FUNCTION_BLOCK FB_DatamanScanner
(*

The function block used to control scanner.

Constructor: 		Patryk Panylo
Company:		E. Riexinger GmbH
Date:			24.01.2019
Version:			1.00

Date:			Revision:		Who:				Comment
dd.mm.yyyy		x.xx			Initials			comment

*)
VAR_INPUT
	(* Input variables / Eingang Variablen *)
	sSrvNetID				:T_AmsNetID	:= '';						(* TwinCAT TCP/IP server network address *)
	sRemoteHost				:T_IPv4Addr := '192.168.10.1';			(* Server network address *)
	nRemotePort				:UDINT := 23;							(* Server port number *)
	bEnable					:BOOL := FALSE;							(* TRUE => enable client data exchange, FALSE => disable *)
	bReset					:BOOL := FALSE;							(* Confirm alarm *)
	bExecute 				:BOOL := FALSE;							(* Send execute command *)
	bLoggerEn				:BOOL := FALSE;							(* TRUE => Enable log message output, FALSE => Disable *)
	sSndMsg					:T_MaxString := 'BEEP 2 2';				(* Send command is an ASCII typable string possibly followed by data. *)
	sPrefix					:STRING := '||>';						(* Send command prefix *)
	sSuffix					:STRING := '$R$N';						(* Send/Receive command suffix *)	
	sDelimiter				:STRING := '';							(* Delimiter (null) *)
	tReceiveTimeout			:TIME := T#100MS;						(* Recive time the which the answer is expected to come *)	
END_VAR
VAR_OUTPUT
	(* Output variables / Ausgang Variablen *)
	sRcvMsg					:T_MaxString := '';						(* Receive an ASCII typable string data. *)										
	arsRcvMsg				:ARRAY[1..GVL_TCPIP.RECEIVE_MESSAGE_MAX] OF T_MaxString;			(* Get message of received an ASCII typable string data. *)
	bConnected				:BOOL := FALSE;							(* TCP/IP connection state connected *)
	bDisconnected			:BOOL := FALSE;							(* TCP/IP connection state disconnected *)
	bRcvDataValid			:BOOL := FALSE;							(* Recive data valid *)	
	bNoDataRcv 				:BOOL := FALSE;							(* No data receive *)	
	bError					:BOOL := FALSE;							(* Program error *)
	bErrorInit				:BOOL := FALSE;							(* Program error initialize *)				
END_VAR
VAR_IN_OUT
	(* Input Output variables / Ausgang Variablen *)

END_VAR
VAR
	(* Enummerations *)
	
	(* Variables *)	
	bInitialize				:BOOL := TRUE;
	
	(* References *)

	(* Interfaces *)

	(* Instances *)
	fbCloseAll				:FB_SocketCloseAll;						(* Close all connection handles (TCP/IP and UDP sockets) that were opened by a PLC runtime system.  *)
	fbConnection			:FB_ClientASCIConnection;				(* Client data exchange control function block. *)
	fbSendMsg 				:FB_ClientSendMsg;						(* Client send cyclic message strings. *)
	fbReceiveMsg 			:FB_ClientReceiveMsg;					(* Client received message strings. *)
	fbLogger 				:FB_ClientLogger;						(* Client get log/error messages from log fifo. *)
	fbTx 					:FB_FrameFifo;							(* Tx fifo *)
	fbRx 					:FB_FrameFifo;							(* Rx fifo *)
	fbLog					:FB_LogFifo;							(* Log/debug/error fifo *)
	fbInitialize			:FB_SignalHandlingDelay;				(* Connection initialize delay *)
	
END_VAR


(* On PLC reset or program download close all old (opened) connections *)
fbInitialize(
	bEnable := TRUE, 
	bIn := bInitialize, 
	tDelay := T#2S
);

fbCloseAll(
	sSrvNetID := sSrvNetID, 
	bExecute := bInitialize 
);

IF fbCloseAll.bBusy 
   OR fbCloseAll.bError 
THEN
	bErrorInit := fbInitialize.bOut;
	RETURN;
ELSE
	bErrorInit := FALSE;
	bInitialize := FALSE;
END_IF

(* Establish connection and data exchange *)
fbConnection(
	bEnable := bEnable, 
	bReset := bReset, 
	bFullDuplex := FALSE, 
	sSrvNetID := sSrvNetID,
	sRemoteHost := sRemoteHost, 
	udnRemotePort := nRemotePort,
	tReconnect := T#45S,
	tReceiveTimeout := tReceiveTimeout,
	bLoggerEn := bLoggerEn, 
	sDelimiter := sDelimiter, 
	sPrefix := 'CLIENT::',
	fbTx := fbTx, 
	fbRx := fbRx, 
	fbLoggger := fbLog, 
	bConnected => bConnected,
	bDisconnected => bDisconnected,
	bRcvDataValid => bRcvDataValid,
	bNoDataRcv => bNoDataRcv,	
	bError => bError
);

(* Send message *)	
fbSendMsg(
	bEnable := bConnected,
	bExecute := bExecute, 
	sMsg := sSndMsg, 
	sPrefix := sPrefix, 
	sSuffix := sSuffix, 
	fbTx := fbTx, 
	fbLoggger := fbLog,
	arsMsg := arsRcvMsg
);

(* Receive message *)	
fbReceiveMsg(
	bEnable := bConnected,
	sSuffix := sSuffix,
	fbRx := fbRx,
	sMsg => sRcvMsg,
	arsMsg := arsRcvMsg
);

(* Log message *)	
fbLogger(
	bEnable := bConnected,
	fbLoggger := fbLog
);

END_FUNCTION_BLOCK

(* stored: Version 1.1.0.1, ProductVersion 3.1.4024.15
   POU FB_DatamanScanner: Id {cff0f39e-88ef-4552-baeb-6b4437f4a8f6}, SpecialFunc None *)
